FUNCTION_BLOCK FB_Ausblasen
VAR_INPUT
END_VAR
VAR_OUTPUT
END_VAR
VAR
tonBlow : TON;
END_VAR

tonBlow(IN := GVL_IO.xAuswerferBereit, PT := T#1S);

GVL_IO.xVentilAusblasenAS := GVL_IO.xAuswerferBereit AND NOT tonBlow.Q;
GVL_IO.xVentilAusblasenGS := NOT GVL_IO.xVentilAusblasenAS;

END_FUNCTION_BLOCK

(* stored: Version 1.1.0.1
   POU FB_Ausblasen: Id {afabcb07-bafc-4fff-915f-45a470bd8161}, SpecialFunc None *)
